(* IEC 61131-3 sources: rusty/tests/lit/cfc/execution_control/enable_chain, 4 files *)

(* ---- main.st ---- *)
FUNCTION main : DINT
    // Both gates FALSE: no gated block ever ran, the ungated ones compute
    // from the defaults, so zeros flow through the whole chain.
    enable_chain();
    // CHECK: idle: counter = 0, d1 = 0, result = 0
    printf('idle: counter = %d, d1 = %d, result = %d$N', enable_chain.c.out, enable_chain.d1.out, enable_chain.result);

    // Both gates TRUE, in sync: 5 accumulates, then (5 * 2 + 1) * 2 = 22.
    enable_chain.g1 := TRUE;
    enable_chain.g2 := TRUE;
    enable_chain();
    // CHECK: sync-on: counter = 5, d1 = 10, result = 22
    printf('sync-on: counter = %d, d1 = %d, result = %d$N', enable_chain.c.out, enable_chain.d1.out, enable_chain.result);

    // Out of sync, head runs and tail holds: the counter advances to 10 and
    // the ungated d1 tracks it to 20, but addOne is frozen at 11, so the
    // tail keeps producing 22; a broken gate would print 42 here.
    enable_chain.g2 := FALSE;
    enable_chain();
    // CHECK: desync-head: counter = 10, d1 = 20, result = 22
    printf('desync-head: counter = %d, d1 = %d, result = %d$N', enable_chain.c.out, enable_chain.d1.out, enable_chain.result);

    // Out of sync the other way, head holds and tail runs: the counter keeps
    // its buffered 10 although seed changed, and the tail recomputes
    // (10 * 2 + 1) * 2 = 42 from that buffer.
    enable_chain.g1 := FALSE;
    enable_chain.g2 := TRUE;
    enable_chain.seed := 100;
    enable_chain();
    // CHECK: desync-tail: counter = 10, d1 = 20, result = 42
    printf('desync-tail: counter = %d, d1 = %d, result = %d$N', enable_chain.c.out, enable_chain.d1.out, enable_chain.result);

    // Both gates FALSE again: everything holds.
    enable_chain.g2 := FALSE;
    enable_chain();
    // CHECK: sync-off: counter = 10, d1 = 20, result = 42
    printf('sync-off: counter = %d, d1 = %d, result = %d$N', enable_chain.c.out, enable_chain.d1.out, enable_chain.result);

    // Both gates TRUE again: the new seed lands, (110 * 2 + 1) * 2 = 442.
    enable_chain.g1 := TRUE;
    enable_chain.g2 := TRUE;
    enable_chain();
    // CHECK: resync: counter = 110, d1 = 220, result = 442
    printf('resync: counter = %d, d1 = %d, result = %d$N', enable_chain.c.out, enable_chain.d1.out, enable_chain.result);
END_FUNCTION

(* ---- addOne.st ---- *)
FUNCTION_BLOCK addOne
VAR_INPUT
    in : DINT;
END_VAR
VAR_OUTPUT
    out : DINT;
END_VAR
    out := in + 1;
END_FUNCTION_BLOCK

(* ---- counter.st ---- *)
FUNCTION_BLOCK counter
VAR_INPUT
    in : DINT;
END_VAR
VAR_OUTPUT
    out : DINT;
END_VAR
    out := out + in;
END_FUNCTION_BLOCK

(* ---- doubler.st ---- *)
FUNCTION_BLOCK doubler
VAR_INPUT
    in : DINT;
END_VAR
VAR_OUTPUT
    out : DINT;
END_VAR
    out := in * 2;
END_FUNCTION_BLOCK
